(* Logix 5000 project; controller SigmaAldrich vendor 1 type 14 code 77 rev 15.4; software revision 15.02; part 2 of 3 *)
(* tags used below, declared in another part *)
   Airlock_N1009_Delay_Tmr : TIMER;
   Airlock_N1009_E_Stop_OSR : BOOL;
   Airlock_N1009_Violation_MDI_Bit : BOOL;
   Airlock_N1009_Violation_MDI_OSR : BOOL;
   Airlock_N1011_E_Stop_OSR : BOOL;
   Airlock_N1011_Violation_MDI_Bit : BOOL;
   Airlock_N1011_Violation_MDI_OSR : BOOL;
   Airlock_N1012_Violation_MDI_Bit : BOOL;
   Airlock_N1012_Violation_MDI_OSR : BOOL;
   Airlock_N1043_E_Stop_OSR : BOOL;
   Airlock_N1043_Violation_MDI_Bit : BOOL;
   Airlock_N1043_Violation_MDI_OSR : BOOL;
   Airlock_N1044_E_Stop_OSR : BOOL;
   Airlock_N1044_Violation_MDI_Bit : BOOL;
   Airlock_N1044_Violation_MDI_OSR : BOOL;
   Airlock_N1052_E_Stop_OSR : BOOL;
   Airlock_N1052_Violation_MDI_Bit : BOOL;
   Airlock_N1052_Violation_MDI_OSR : BOOL;
   Airlock_N1065_E_Stop_OSR : BOOL;
   Airlock_N1065_Violation_MDI_Bit : BOOL;
   Airlock_N1065_Violation_MDI_OSR : BOOL;
   Airlock_N1066_E_Stop_OSR : BOOL;
   Airlock_N1066_Violation_MDI_Bit : BOOL;
   Airlock_N1066_Violation_MDI_OSR : BOOL;
   Annuciator_Bit_Airlock_N1009 : BOOL;
   Annuciator_Bit_Airlock_N1011 : BOOL;
   Annuciator_Bit_Airlock_N1012 : BOOL;
   Annuciator_Bit_Airlock_N1043 : BOOL;
   Annuciator_Bit_Airlock_N1044 : BOOL;
   Annuciator_Bit_Airlock_N1052 : BOOL;
   Annuciator_Bit_Airlock_N1065 : BOOL;
   Annuciator_Bit_Airlock_N1066 : BOOL;
   Door_N1009A_Timer : TIMER;
   Door_N1009B_Timer : TIMER;
   Door_N1011A_Timer : TIMER;
   Door_N1011B_Timer : TIMER;
   Door_N1012_Timer : TIMER;
   Door_N1043A_Timer : TIMER;
   Door_N1043B_Timer : TIMER;
   Door_N1044A_Timer : TIMER;
   Door_N1044B_Timer : TIMER;
   Door_N1044C_Timer : TIMER;
   Door_N1052A_Timer : TIMER;
   Door_N1052B_Timer : TIMER;
   Door_N1053_Timer : TIMER;
   Door_N1058B_Timer : TIMER;
   Door_N1065A_Timer : TIMER;
   Door_N1065B_Timer : TIMER;
   Door_N1066A_Timer : TIMER;
   Door_N1066B_Timer : TIMER;
   MDI_Violation_N1009_Bit : BOOL;
   MDI_Violation_N1011_Bit : BOOL;
   MDI_Violation_N1012_Bit : BOOL;
   MDI_Violation_N1043_Bit : BOOL;
   MDI_Violation_N1044_Bit : BOOL;
   MDI_Violation_N1052_Bit : BOOL;
   MDI_Violation_N1065_Bit : BOOL;
   MDI_Violation_N1066_Bit : BOOL;
   N1008_Emergency_Release_Latch : BOOL;
   N1009_Airlock_Latch : BOOL;
   N1009_Emergency_Release_Latch : BOOL;
   N1011_Airlock_Latch : BOOL;
   N1011_Emergency_Release_Latch : BOOL;
   N1012_Airlock_Latch : BOOL;
   N1012_Emergency_Release_Latch : BOOL;
   N1043_Airlock_Latch : BOOL;
   N1043_Emergency_Release_Latch : BOOL;
   N1044_Airlock_Latch : BOOL;
   N1044_Emergency_Release_Latch : BOOL;
   N1044A_Door_Latch_Bit : BOOL;
   N1052_Airlock_Latch : BOOL;
   N1052_Emergency_Release_Latch : BOOL;
   N1052A_Door_Latch_Bit : BOOL;
   N1065_Airlock_Latch : BOOL;
   N1065_Emergency_Release_Latch : BOOL;
   N1066_Airlock_Latch : BOOL;
   N1066_Emergency_Release_Latch : BOOL;
(* MainProgram, continued *)

ROUTINE DI07_N1009   (* ladder *)
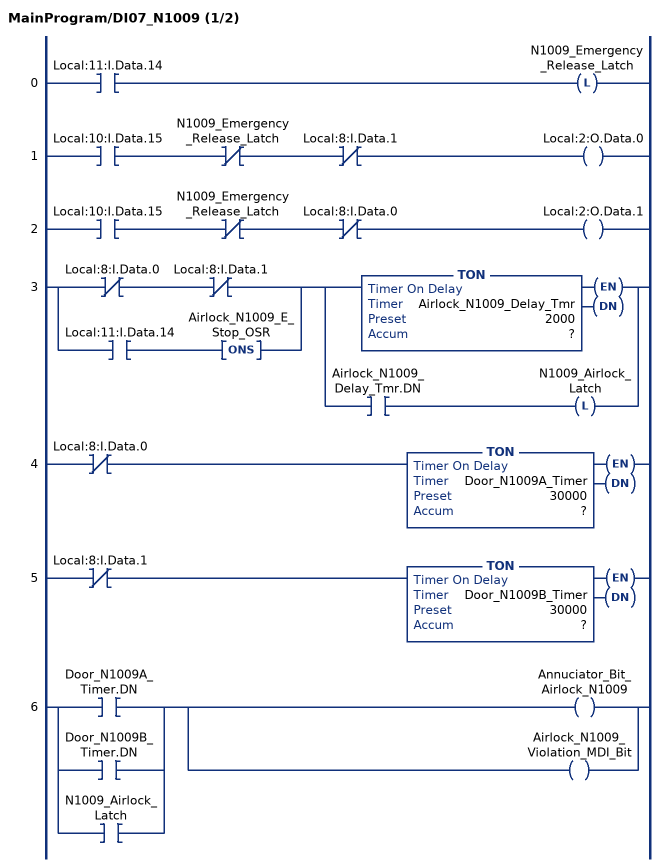
   0: XIC(Local:11:I.Data.14)OTL(N1009_Emergency_Release_Latch);
   1: XIC(Local:10:I.Data.15)XIO(N1009_Emergency_Release_Latch)XIO(Local:8:I.Data.1)OTE(Local:2:O.Data.0);
   2: XIC(Local:10:I.Data.15)XIO(N1009_Emergency_Release_Latch)XIO(Local:8:I.Data.0)OTE(Local:2:O.Data.1);
   3: [XIO(Local:8:I.Data.0) XIO(Local:8:I.Data.1) ,XIC(Local:11:I.Data.14) ONS(Airlock_N1009_E_Stop_OSR) ][TON(Airlock_N1009_Delay_Tmr,?,?) ,XIC(Airlock_N1009_Delay_Tmr.DN) OTL(N1009_Airlock_Latch) ];
   4: XIO(Local:8:I.Data.0)TON(Door_N1009A_Timer,?,?);
   5: XIO(Local:8:I.Data.1)TON(Door_N1009B_Timer,?,?);
   6: [XIC(Door_N1009A_Timer.DN) ,XIC(Door_N1009B_Timer.DN) ,XIC(N1009_Airlock_Latch) ][OTE(Annuciator_Bit_Airlock_N1009) ,OTE(Airlock_N1009_Violation_MDI_Bit) ];
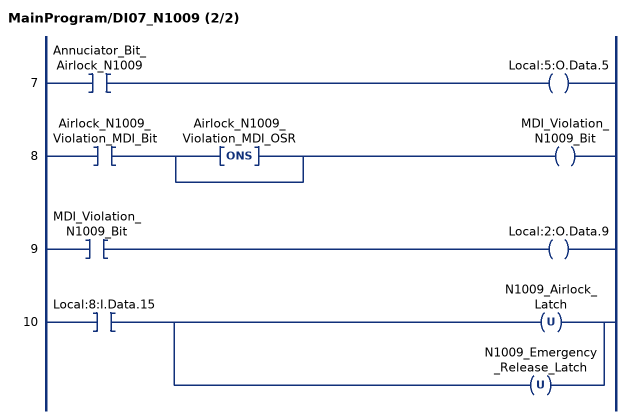
   7: XIC(Annuciator_Bit_Airlock_N1009)OTE(Local:5:O.Data.5);
   8: XIC(Airlock_N1009_Violation_MDI_Bit)[ONS(Airlock_N1009_Violation_MDI_OSR) ,]OTE(MDI_Violation_N1009_Bit);
   9: XIC(MDI_Violation_N1009_Bit)OTE(Local:2:O.Data.9);
   10: XIC(Local:8:I.Data.15)[OTU(N1009_Airlock_Latch) ,OTU(N1009_Emergency_Release_Latch) ];
END_ROUTINE

ROUTINE DI08_N1011   (* ladder *)
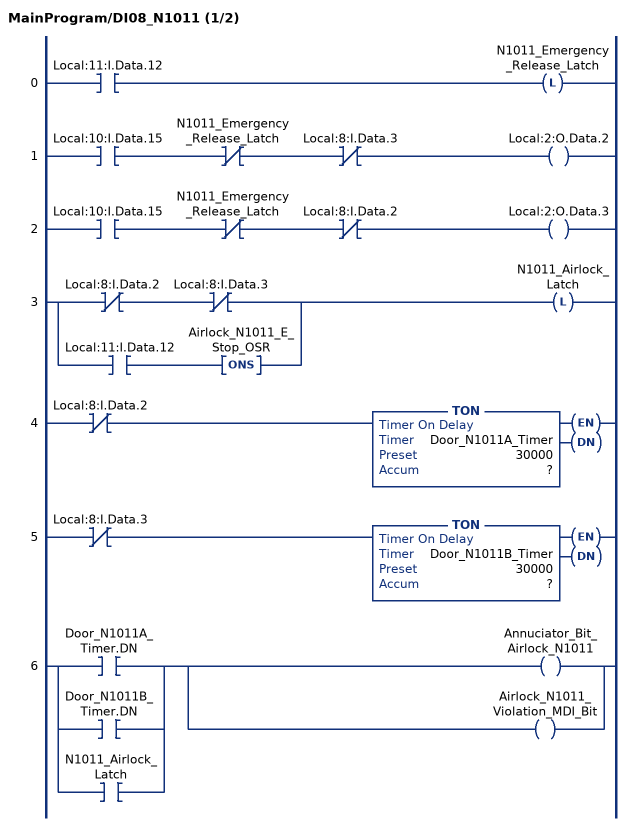
   0: XIC(Local:11:I.Data.12)OTL(N1011_Emergency_Release_Latch);
   1: XIC(Local:10:I.Data.15)XIO(N1011_Emergency_Release_Latch)XIO(Local:8:I.Data.3)OTE(Local:2:O.Data.2);
   2: XIC(Local:10:I.Data.15)XIO(N1011_Emergency_Release_Latch)XIO(Local:8:I.Data.2)OTE(Local:2:O.Data.3);
   3: [XIO(Local:8:I.Data.2) XIO(Local:8:I.Data.3) ,XIC(Local:11:I.Data.12) ONS(Airlock_N1011_E_Stop_OSR) ]OTL(N1011_Airlock_Latch);
   4: XIO(Local:8:I.Data.2)TON(Door_N1011A_Timer,?,?);
   5: XIO(Local:8:I.Data.3)TON(Door_N1011B_Timer,?,?);
   6: [XIC(Door_N1011A_Timer.DN) ,XIC(Door_N1011B_Timer.DN) ,XIC(N1011_Airlock_Latch) ][OTE(Annuciator_Bit_Airlock_N1011) ,OTE(Airlock_N1011_Violation_MDI_Bit) ];
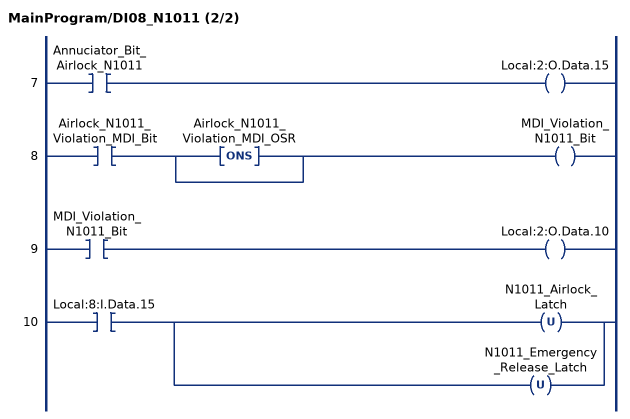
   7: XIC(Annuciator_Bit_Airlock_N1011)OTE(Local:2:O.Data.15);
   8: XIC(Airlock_N1011_Violation_MDI_Bit)[ONS(Airlock_N1011_Violation_MDI_OSR) ,]OTE(MDI_Violation_N1011_Bit);
   9: XIC(MDI_Violation_N1011_Bit)OTE(Local:2:O.Data.10);
   10: XIC(Local:8:I.Data.15)[OTU(N1011_Airlock_Latch) ,OTU(N1011_Emergency_Release_Latch) ];
END_ROUTINE

ROUTINE DI09_N1012   (* ladder *)
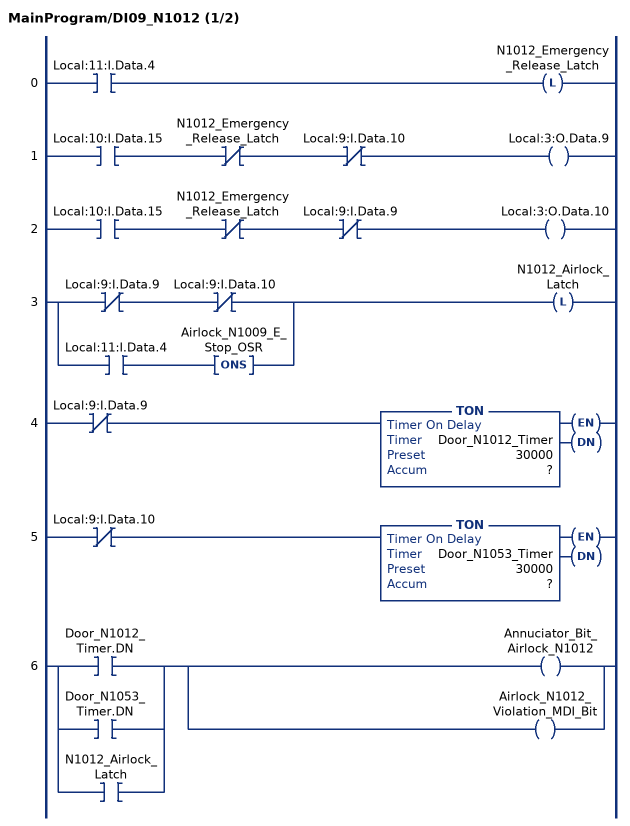
   0: XIC(Local:11:I.Data.4)OTL(N1012_Emergency_Release_Latch);
   1: XIC(Local:10:I.Data.15)XIO(N1012_Emergency_Release_Latch)XIO(Local:9:I.Data.10)OTE(Local:3:O.Data.9);
   2: XIC(Local:10:I.Data.15)XIO(N1012_Emergency_Release_Latch)XIO(Local:9:I.Data.9)OTE(Local:3:O.Data.10);
   3: [XIO(Local:9:I.Data.9) XIO(Local:9:I.Data.10) ,XIC(Local:11:I.Data.4) ONS(Airlock_N1009_E_Stop_OSR) ]OTL(N1012_Airlock_Latch);
   4: XIO(Local:9:I.Data.9)TON(Door_N1012_Timer,?,?);
   5: XIO(Local:9:I.Data.10)TON(Door_N1053_Timer,?,?);
   6: [XIC(Door_N1012_Timer.DN) ,XIC(Door_N1053_Timer.DN) ,XIC(N1012_Airlock_Latch) ][OTE(Annuciator_Bit_Airlock_N1012) ,OTE(Airlock_N1012_Violation_MDI_Bit) ];
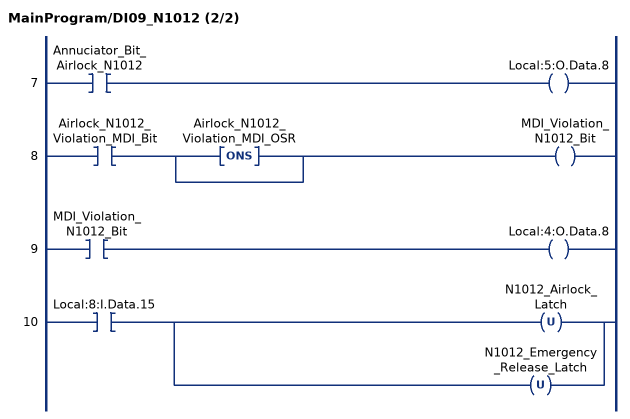
   7: XIC(Annuciator_Bit_Airlock_N1012)OTE(Local:5:O.Data.8);
   8: XIC(Airlock_N1012_Violation_MDI_Bit)[ONS(Airlock_N1012_Violation_MDI_OSR) ,]OTE(MDI_Violation_N1012_Bit);
   9: XIC(MDI_Violation_N1012_Bit)OTE(Local:4:O.Data.8);
   10: XIC(Local:8:I.Data.15)[OTU(N1012_Airlock_Latch) ,OTU(N1012_Emergency_Release_Latch) ];
END_ROUTINE

ROUTINE DI10_N1043   (* ladder *)
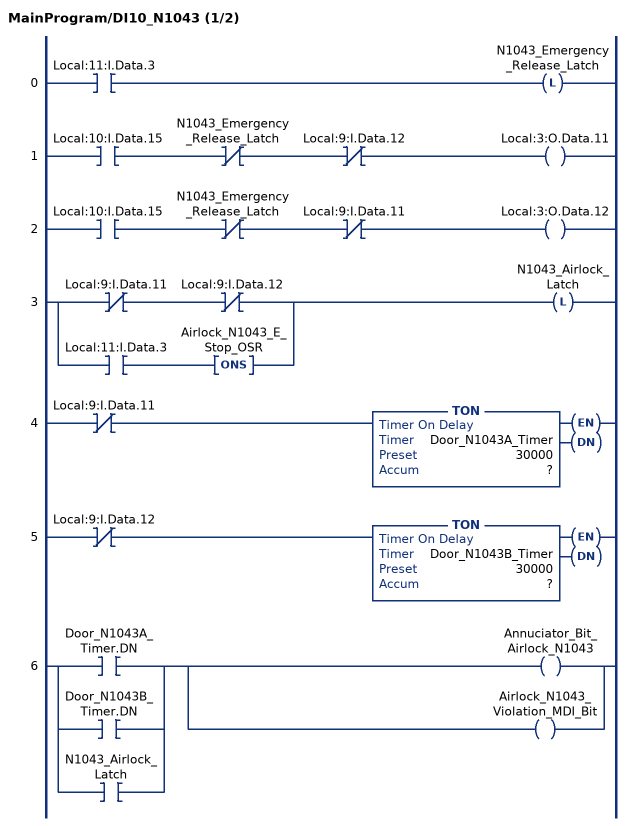
   0: XIC(Local:11:I.Data.3)OTL(N1043_Emergency_Release_Latch);
   1: XIC(Local:10:I.Data.15)XIO(N1043_Emergency_Release_Latch)XIO(Local:9:I.Data.12)OTE(Local:3:O.Data.11);
   2: XIC(Local:10:I.Data.15)XIO(N1043_Emergency_Release_Latch)XIO(Local:9:I.Data.11)OTE(Local:3:O.Data.12);
   3: [XIO(Local:9:I.Data.11) XIO(Local:9:I.Data.12) ,XIC(Local:11:I.Data.3) ONS(Airlock_N1043_E_Stop_OSR) ]OTL(N1043_Airlock_Latch);
   4: XIO(Local:9:I.Data.11)TON(Door_N1043A_Timer,?,?);
   5: XIO(Local:9:I.Data.12)TON(Door_N1043B_Timer,?,?);
   6: [XIC(Door_N1043A_Timer.DN) ,XIC(Door_N1043B_Timer.DN) ,XIC(N1043_Airlock_Latch) ][OTE(Annuciator_Bit_Airlock_N1043) ,OTE(Airlock_N1043_Violation_MDI_Bit) ];
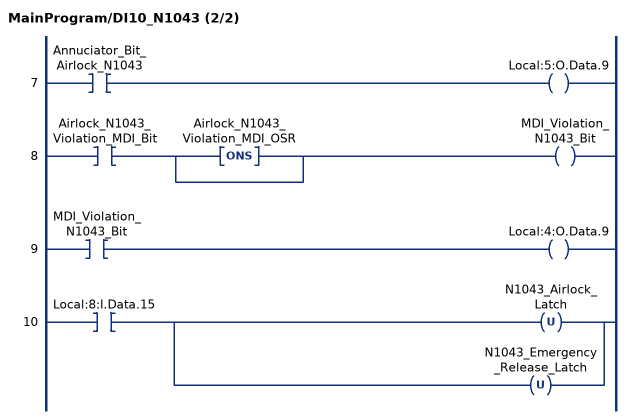
   7: XIC(Annuciator_Bit_Airlock_N1043)OTE(Local:5:O.Data.9);
   8: XIC(Airlock_N1043_Violation_MDI_Bit)[ONS(Airlock_N1043_Violation_MDI_OSR) ,]OTE(MDI_Violation_N1043_Bit);
   9: XIC(MDI_Violation_N1043_Bit)OTE(Local:4:O.Data.9);
   10: XIC(Local:8:I.Data.15)[OTU(N1043_Airlock_Latch) ,OTU(N1043_Emergency_Release_Latch) ];
END_ROUTINE

ROUTINE DI11_N1044   (* ladder *)
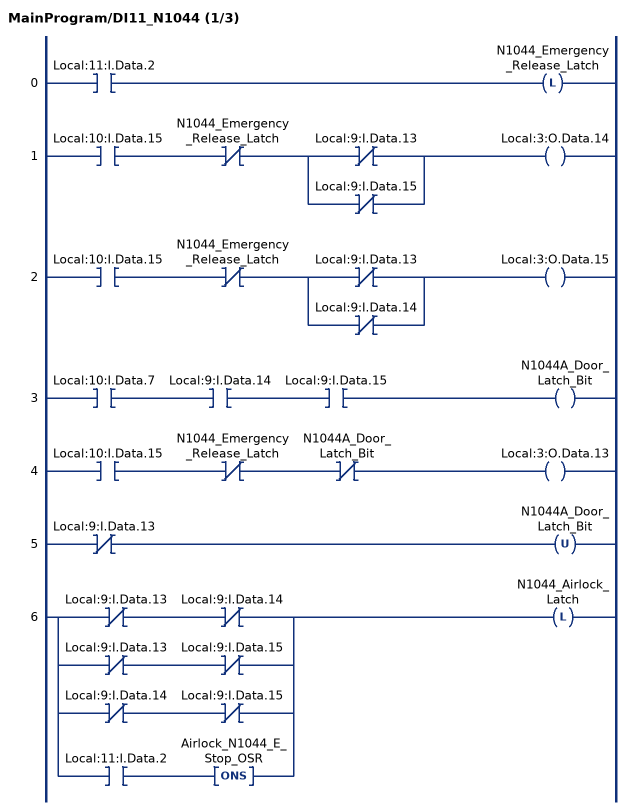
   0: XIC(Local:11:I.Data.2)OTL(N1044_Emergency_Release_Latch);
   1: XIC(Local:10:I.Data.15)XIO(N1044_Emergency_Release_Latch)[XIO(Local:9:I.Data.13) ,XIO(Local:9:I.Data.15) ]OTE(Local:3:O.Data.14);
   2: XIC(Local:10:I.Data.15)XIO(N1044_Emergency_Release_Latch)[XIO(Local:9:I.Data.13) ,XIO(Local:9:I.Data.14) ]OTE(Local:3:O.Data.15);
   3: XIC(Local:10:I.Data.7)XIC(Local:9:I.Data.14)XIC(Local:9:I.Data.15)OTE(N1044A_Door_Latch_Bit);
   4: XIC(Local:10:I.Data.15)XIO(N1044_Emergency_Release_Latch)XIO(N1044A_Door_Latch_Bit)OTE(Local:3:O.Data.13);
   5: XIO(Local:9:I.Data.13)OTU(N1044A_Door_Latch_Bit);
   6: [XIO(Local:9:I.Data.13) XIO(Local:9:I.Data.14) ,XIO(Local:9:I.Data.13) XIO(Local:9:I.Data.15) ,XIO(Local:9:I.Data.14) XIO(Local:9:I.Data.15) ,XIC(Local:11:I.Data.2) ONS(Airlock_N1044_E_Stop_OSR) ]OTL(N1044_Airlock_Latch);
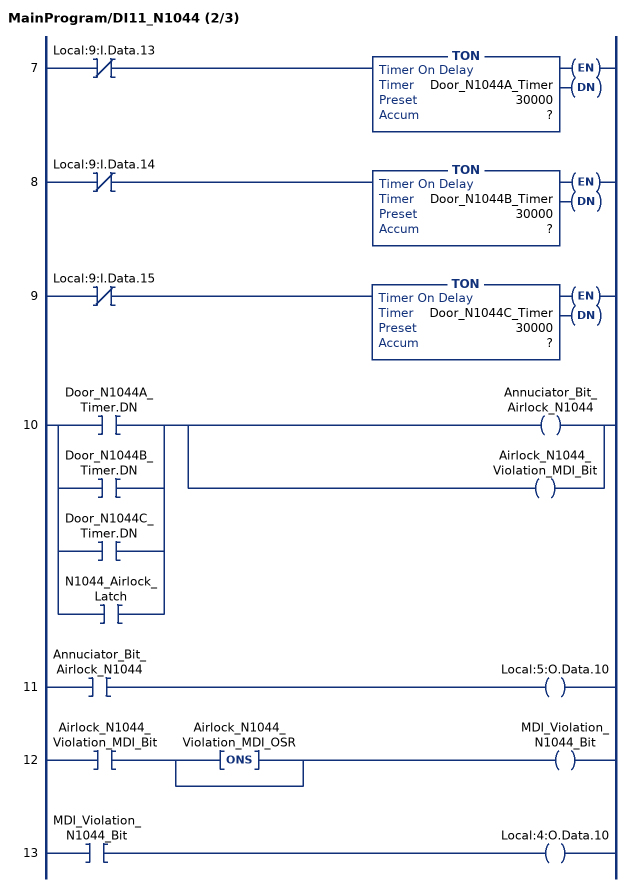
   7: XIO(Local:9:I.Data.13)TON(Door_N1044A_Timer,?,?);
   8: XIO(Local:9:I.Data.14)TON(Door_N1044B_Timer,?,?);
   9: XIO(Local:9:I.Data.15)TON(Door_N1044C_Timer,?,?);
   10: [XIC(Door_N1044A_Timer.DN) ,XIC(Door_N1044B_Timer.DN) ,XIC(Door_N1044C_Timer.DN) ,XIC(N1044_Airlock_Latch) ][OTE(Annuciator_Bit_Airlock_N1044) ,OTE(Airlock_N1044_Violation_MDI_Bit) ];
   11: XIC(Annuciator_Bit_Airlock_N1044)OTE(Local:5:O.Data.10);
   12: XIC(Airlock_N1044_Violation_MDI_Bit)[ONS(Airlock_N1044_Violation_MDI_OSR) ,]OTE(MDI_Violation_N1044_Bit);
   13: XIC(MDI_Violation_N1044_Bit)OTE(Local:4:O.Data.10);
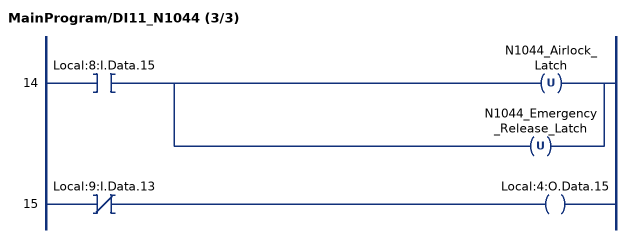
   14: XIC(Local:8:I.Data.15)[OTU(N1044_Airlock_Latch) ,OTU(N1044_Emergency_Release_Latch) ];
   15: XIO(Local:9:I.Data.13)OTE(Local:4:O.Data.15);
END_ROUTINE

ROUTINE DI12_N1052   (* ladder *)
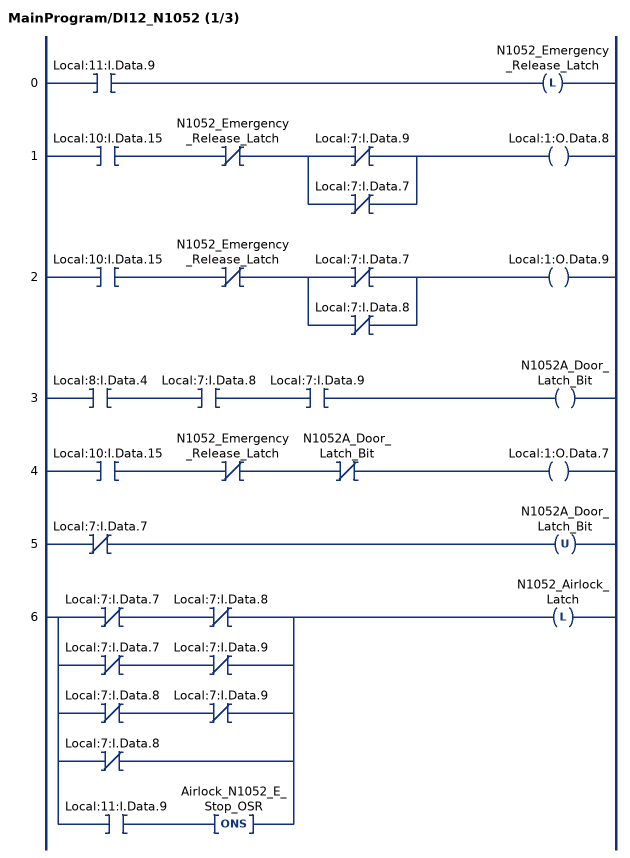
   0: XIC(Local:11:I.Data.9)OTL(N1052_Emergency_Release_Latch);
   1: XIC(Local:10:I.Data.15)XIO(N1052_Emergency_Release_Latch)[XIO(Local:7:I.Data.9) ,XIO(Local:7:I.Data.7) ]OTE(Local:1:O.Data.8);
   2: XIC(Local:10:I.Data.15)XIO(N1052_Emergency_Release_Latch)[XIO(Local:7:I.Data.7) ,XIO(Local:7:I.Data.8) ]OTE(Local:1:O.Data.9);
   3: XIC(Local:8:I.Data.4)XIC(Local:7:I.Data.8)XIC(Local:7:I.Data.9)OTE(N1052A_Door_Latch_Bit);
   4: XIC(Local:10:I.Data.15)XIO(N1052_Emergency_Release_Latch)XIO(N1052A_Door_Latch_Bit)OTE(Local:1:O.Data.7);
   5: XIO(Local:7:I.Data.7)OTU(N1052A_Door_Latch_Bit);
   6: [XIO(Local:7:I.Data.7) XIO(Local:7:I.Data.8) ,XIO(Local:7:I.Data.7) XIO(Local:7:I.Data.9) ,XIO(Local:7:I.Data.8) XIO(Local:7:I.Data.9) ,XIO(Local:7:I.Data.8) ,XIC(Local:11:I.Data.9) ONS(Airlock_N1052_E_Stop_OSR) ]OTL(N1052_Airlock_Latch);
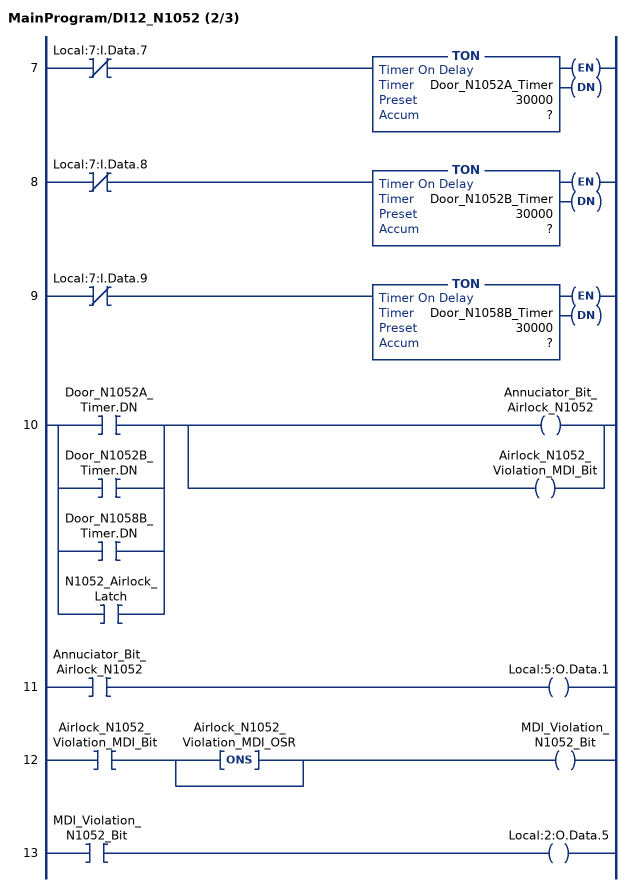
   7: XIO(Local:7:I.Data.7)TON(Door_N1052A_Timer,?,?);
   8: XIO(Local:7:I.Data.8)TON(Door_N1052B_Timer,?,?);
   9: XIO(Local:7:I.Data.9)TON(Door_N1058B_Timer,?,?);
   10: [XIC(Door_N1052A_Timer.DN) ,XIC(Door_N1052B_Timer.DN) ,XIC(Door_N1058B_Timer.DN) ,XIC(N1052_Airlock_Latch) ][OTE(Annuciator_Bit_Airlock_N1052) ,OTE(Airlock_N1052_Violation_MDI_Bit) ];
   11: XIC(Annuciator_Bit_Airlock_N1052)OTE(Local:5:O.Data.1);
   12: XIC(Airlock_N1052_Violation_MDI_Bit)[ONS(Airlock_N1052_Violation_MDI_OSR) ,]OTE(MDI_Violation_N1052_Bit);
   13: XIC(MDI_Violation_N1052_Bit)OTE(Local:2:O.Data.5);
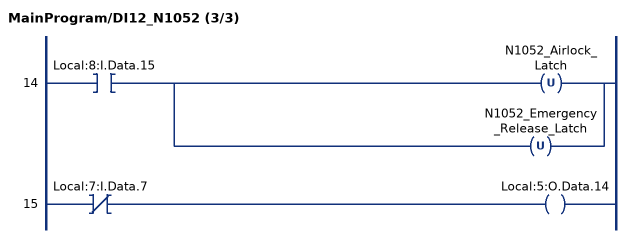
   14: XIC(Local:8:I.Data.15)[OTU(N1052_Airlock_Latch) ,OTU(N1052_Emergency_Release_Latch) ];
   15: XIO(Local:7:I.Data.7)OTE(Local:5:O.Data.14);
END_ROUTINE

ROUTINE DI13_N1065   (* ladder *)
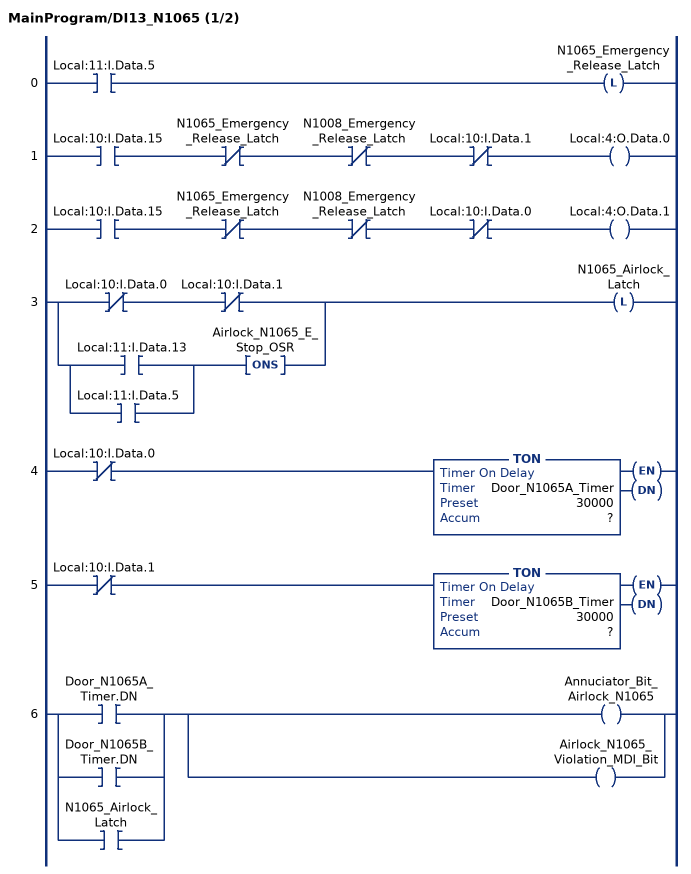
   0: XIC(Local:11:I.Data.5)OTL(N1065_Emergency_Release_Latch);
   1: XIC(Local:10:I.Data.15)XIO(N1065_Emergency_Release_Latch)XIO(N1008_Emergency_Release_Latch)XIO(Local:10:I.Data.1)OTE(Local:4:O.Data.0);
   2: XIC(Local:10:I.Data.15)XIO(N1065_Emergency_Release_Latch)XIO(N1008_Emergency_Release_Latch)XIO(Local:10:I.Data.0)OTE(Local:4:O.Data.1);
   3: [XIO(Local:10:I.Data.0) XIO(Local:10:I.Data.1) ,[XIC(Local:11:I.Data.13) ,XIC(Local:11:I.Data.5) ] ONS(Airlock_N1065_E_Stop_OSR) ]OTL(N1065_Airlock_Latch);
   4: XIO(Local:10:I.Data.0)TON(Door_N1065A_Timer,?,?);
   5: XIO(Local:10:I.Data.1)TON(Door_N1065B_Timer,?,?);
   6: [XIC(Door_N1065A_Timer.DN) ,XIC(Door_N1065B_Timer.DN) ,XIC(N1065_Airlock_Latch) ][OTE(Annuciator_Bit_Airlock_N1065) ,OTE(Airlock_N1065_Violation_MDI_Bit) ];
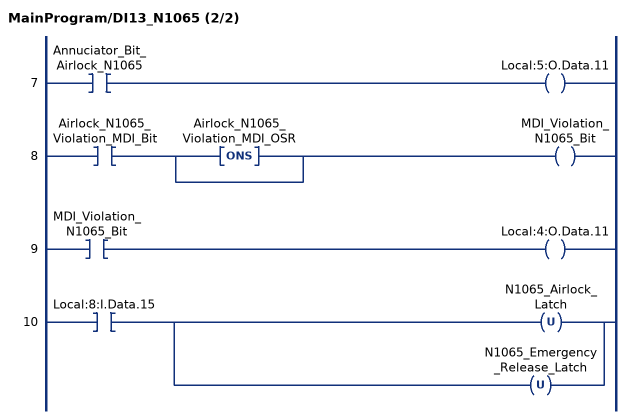
   7: XIC(Annuciator_Bit_Airlock_N1065)OTE(Local:5:O.Data.11);
   8: XIC(Airlock_N1065_Violation_MDI_Bit)[ONS(Airlock_N1065_Violation_MDI_OSR) ,]OTE(MDI_Violation_N1065_Bit);
   9: XIC(MDI_Violation_N1065_Bit)OTE(Local:4:O.Data.11);
   10: XIC(Local:8:I.Data.15)[OTU(N1065_Airlock_Latch) ,OTU(N1065_Emergency_Release_Latch) ];
END_ROUTINE

ROUTINE DI14_N1066   (* ladder *)
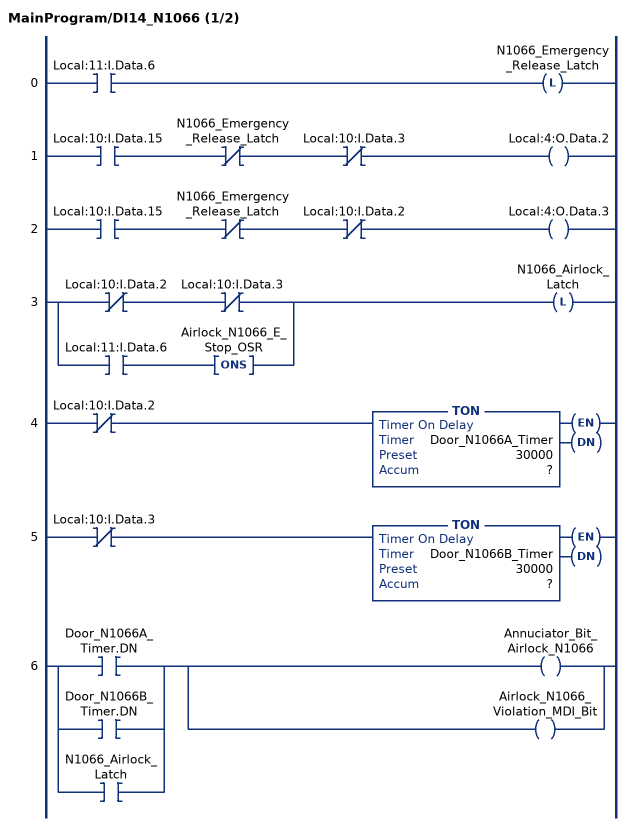
   0: XIC(Local:11:I.Data.6)OTL(N1066_Emergency_Release_Latch);
   1: XIC(Local:10:I.Data.15)XIO(N1066_Emergency_Release_Latch)XIO(Local:10:I.Data.3)OTE(Local:4:O.Data.2);
   2: XIC(Local:10:I.Data.15)XIO(N1066_Emergency_Release_Latch)XIO(Local:10:I.Data.2)OTE(Local:4:O.Data.3);
   3: [XIO(Local:10:I.Data.2) XIO(Local:10:I.Data.3) ,XIC(Local:11:I.Data.6) ONS(Airlock_N1066_E_Stop_OSR) ]OTL(N1066_Airlock_Latch);
   4: XIO(Local:10:I.Data.2)TON(Door_N1066A_Timer,?,?);
   5: XIO(Local:10:I.Data.3)TON(Door_N1066B_Timer,?,?);
   6: [XIC(Door_N1066A_Timer.DN) ,XIC(Door_N1066B_Timer.DN) ,XIC(N1066_Airlock_Latch) ][OTE(Annuciator_Bit_Airlock_N1066) ,OTE(Airlock_N1066_Violation_MDI_Bit) ];
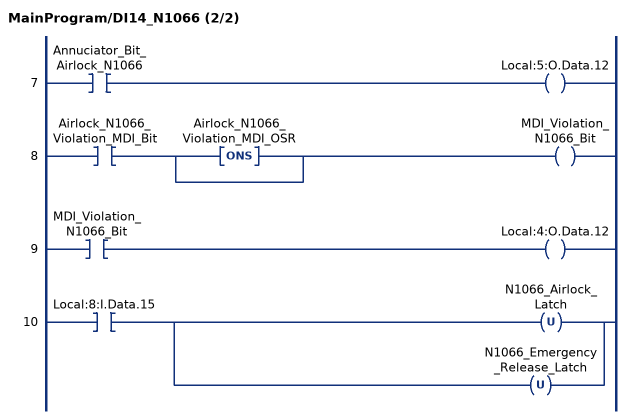
   7: XIC(Annuciator_Bit_Airlock_N1066)OTE(Local:5:O.Data.12);
   8: XIC(Airlock_N1066_Violation_MDI_Bit)[ONS(Airlock_N1066_Violation_MDI_OSR) ,]OTE(MDI_Violation_N1066_Bit);
   9: XIC(MDI_Violation_N1066_Bit)OTE(Local:4:O.Data.12);
   10: XIC(Local:8:I.Data.15)[OTU(N1066_Airlock_Latch) ,OTU(N1066_Emergency_Release_Latch) ];
END_ROUTINE
